(* IEC 61131-3 sources: ironplc/compiler/syntax/tests/fixtures/malformed, 12 files *)

(* ---- mismatched_closers.st ---- *)
FUNCTION_BLOCK Fb
VAR x : INT; END_VAR
x := 1;
END_PROGRAM

FUNCTION f : INT
f := 1;
END_FUNCTION_BLOCK

(* ---- unterminated_method.st ---- *)
FUNCTION_BLOCK Fb
VAR x : INT; END_VAR
METHOD Run : BOOL
    Run := TRUE;
END_FUNCTION_BLOCK

PROGRAM Main
END_PROGRAM

(* ---- bad_type_declarations.st ---- *)
TYPE
    Good : INT := 5;
    Broken : ARRAY[1..] OF INT;
    Colors : (Red, Green, Blue);
    Point : STRUCT
        x : INT;
        y : ;
    END_STRUCT;
END_TYPE

PROGRAM After
END_PROGRAM

(* ---- broken_declarations.st ---- *)
PROGRAM Broken
VAR
	ok : INT;
	missing : ;
	p AT : INT;
	ok2 : INT;
END_VAR
x := f(,);
END_PROGRAM

(* ---- dangling_operator.st ---- *)
PROGRAM P
x := 1 + ;
y := 2;
END_PROGRAM

(* ---- empty_and_missing_parts.st ---- *)
PROGRAM
END_PROGRAM
FUNCTION : INT
END_FUNCTION
FUNCTION g
g := 1;
END_FUNCTION
TYPE END_TYPE
VAR_GLOBAL
    a : INT
    b : INT;
END_VAR

(* ---- missing_end_program.st ---- *)
PROGRAM First
VAR a : INT; END_VAR
a := 1;

PROGRAM Second
VAR b : INT; END_VAR
b := 2;
END_PROGRAM

(* ---- stray_between_programs.st ---- *)
PROGRAM A
END_PROGRAM
???
PROGRAM B
END_PROGRAM

(* ---- stray_end_var.st ---- *)
PROGRAM P
VAR x : INT; END_VAR
END_VAR
x := 1;
IF x > 0 THEN
    x := 2;
END_PROGRAM

(* ---- unknown_character.st ---- *)
PROGRAM P
x := 1 ? 2;
END_PROGRAM

(* ---- unterminated_comment.st ---- *)
PROGRAM P
(* never closed
END_PROGRAM

(* ---- unterminated_var_block.st ---- *)
PROGRAM Open
VAR
    a : INT;
    b : BOOL;
x := 1;
END_PROGRAM

PROGRAM Next
VAR c : INT; END_VAR
c := 2;
END_PROGRAM
